(* IEC 61131-3 sources: stonehenge-public/apps/core/stonehenge-safety-plc/pous/programs, 1 file *)

(* ---- main.st ---- *)
PROGRAM main
  VAR
    SafetyGlobal : FB_GlobalSafety;
    Gun1Safety : FB_GunSafety;
    Gun2Safety : FB_GunSafety;
    Gun3Safety : FB_GunSafety;
    Gun4Safety : FB_GunSafety;
    Gun5Safety : FB_GunSafety;
    Gun6Safety : FB_GunSafety;
    Gun7Safety : FB_GunSafety;
    Gun8Safety : FB_GunSafety;
    CONTROL_VERSION_REQUEST : INT AT %MW0 := 0;
    GLOBAL_ENABLE : INT AT %MW1 := 0;
    EMERGENCY_STOP : INT AT %MW2 := 0;
    GLOBAL_MAINTENANCE_MODE : INT AT %MW3 := 0;
    SAFETY_RESET_REQUEST : INT AT %MW4 := 0;
    TEST_FAULT_REQUEST : INT AT %MW5 := 0;
    INPUT_RESERVED_6 : INT AT %MW6 := 0;
    INPUT_RESERVED_7 : INT AT %MW7 := 0;
    GUN1_ENABLED : INT AT %MW16 := 0;
    GUN1_MAINTENANCE_INHIBIT : INT AT %MW17 := 0;
    GUN1_EXTERNAL_INHIBIT : INT AT %MW18 := 0;
    GUN1_INPUT_RESERVED : INT AT %MW19 := 0;
    GUN2_ENABLED : INT AT %MW20 := 0;
    GUN2_MAINTENANCE_INHIBIT : INT AT %MW21 := 0;
    GUN2_EXTERNAL_INHIBIT : INT AT %MW22 := 0;
    GUN2_INPUT_RESERVED : INT AT %MW23 := 0;
    GUN3_ENABLED : INT AT %MW24 := 0;
    GUN3_MAINTENANCE_INHIBIT : INT AT %MW25 := 0;
    GUN3_EXTERNAL_INHIBIT : INT AT %MW26 := 0;
    GUN3_INPUT_RESERVED : INT AT %MW27 := 0;
    GUN4_ENABLED : INT AT %MW28 := 0;
    GUN4_MAINTENANCE_INHIBIT : INT AT %MW29 := 0;
    GUN4_EXTERNAL_INHIBIT : INT AT %MW30 := 0;
    GUN4_INPUT_RESERVED : INT AT %MW31 := 0;
    GUN5_ENABLED : INT AT %MW32 := 0;
    GUN5_MAINTENANCE_INHIBIT : INT AT %MW33 := 0;
    GUN5_EXTERNAL_INHIBIT : INT AT %MW34 := 0;
    GUN5_INPUT_RESERVED : INT AT %MW35 := 0;
    GUN6_ENABLED : INT AT %MW36 := 0;
    GUN6_MAINTENANCE_INHIBIT : INT AT %MW37 := 0;
    GUN6_EXTERNAL_INHIBIT : INT AT %MW38 := 0;
    GUN6_INPUT_RESERVED : INT AT %MW39 := 0;
    GUN7_ENABLED : INT AT %MW40 := 0;
    GUN7_MAINTENANCE_INHIBIT : INT AT %MW41 := 0;
    GUN7_EXTERNAL_INHIBIT : INT AT %MW42 := 0;
    GUN7_INPUT_RESERVED : INT AT %MW43 := 0;
    GUN8_ENABLED : INT AT %MW44 := 0;
    GUN8_MAINTENANCE_INHIBIT : INT AT %MW45 := 0;
    GUN8_EXTERNAL_INHIBIT : INT AT %MW46 := 0;
    GUN8_INPUT_RESERVED : INT AT %MW47 := 0;
    SAFETY_SCHEMA_VERSION : INT AT %QW0 := 0;
    SAFETY_HEARTBEAT_COUNTER : INT AT %QW1 := 0;
    SAFETY_STATE : INT AT %QW2 := 0;
    SAFETY_READY : INT AT %QW3 := 0;
    GLOBAL_FIRE_PERMISSIVE : INT AT %QW4 := 0;
    GLOBAL_INHIBIT_ACTIVE : INT AT %QW5 := 0;
    GLOBAL_INHIBIT_REASON : INT AT %QW6 := 0;
    SAFETY_FAULT_ACTIVE : INT AT %QW7 := 0;
    SAFETY_FAULT_CODE : INT AT %QW8 := 0;
    RESET_REQUIRED : INT AT %QW9 := 0;
    EMERGENCY_STOP_ACTIVE : INT AT %QW10 := 0;
    MAINTENANCE_MODE_ACTIVE : INT AT %QW11 := 0;
    STATUS_RESERVED_12 : INT AT %QW12 := 0;
    STATUS_RESERVED_13 : INT AT %QW13 := 0;
    STATUS_RESERVED_14 : INT AT %QW14 := 0;
    STATUS_RESERVED_15 : INT AT %QW15 := 0;
    GUN1_FIRE_PERMISSIVE : INT AT %QW16 := 0;
    GUN1_INHIBIT_ACTIVE : INT AT %QW17 := 0;
    GUN1_INHIBIT_REASON : INT AT %QW18 := 0;
    GUN1_ENABLED_STATUS : INT AT %QW19 := 0;
    GUN1_MAINTENANCE_INHIBIT_STATUS : INT AT %QW20 := 0;
    GUN1_EXTERNAL_INHIBIT_STATUS : INT AT %QW21 := 0;
    GUN1_STATUS_RESERVED_A : INT AT %QW22 := 0;
    GUN1_STATUS_RESERVED_B : INT AT %QW23 := 0;
    GUN2_FIRE_PERMISSIVE : INT AT %QW24 := 0;
    GUN2_INHIBIT_ACTIVE : INT AT %QW25 := 0;
    GUN2_INHIBIT_REASON : INT AT %QW26 := 0;
    GUN2_ENABLED_STATUS : INT AT %QW27 := 0;
    GUN2_MAINTENANCE_INHIBIT_STATUS : INT AT %QW28 := 0;
    GUN2_EXTERNAL_INHIBIT_STATUS : INT AT %QW29 := 0;
    GUN2_STATUS_RESERVED_A : INT AT %QW30 := 0;
    GUN2_STATUS_RESERVED_B : INT AT %QW31 := 0;
    GUN3_FIRE_PERMISSIVE : INT AT %QW32 := 0;
    GUN3_INHIBIT_ACTIVE : INT AT %QW33 := 0;
    GUN3_INHIBIT_REASON : INT AT %QW34 := 0;
    GUN3_ENABLED_STATUS : INT AT %QW35 := 0;
    GUN3_MAINTENANCE_INHIBIT_STATUS : INT AT %QW36 := 0;
    GUN3_EXTERNAL_INHIBIT_STATUS : INT AT %QW37 := 0;
    GUN3_STATUS_RESERVED_A : INT AT %QW38 := 0;
    GUN3_STATUS_RESERVED_B : INT AT %QW39 := 0;
    GUN4_FIRE_PERMISSIVE : INT AT %QW40 := 0;
    GUN4_INHIBIT_ACTIVE : INT AT %QW41 := 0;
    GUN4_INHIBIT_REASON : INT AT %QW42 := 0;
    GUN4_ENABLED_STATUS : INT AT %QW43 := 0;
    GUN4_MAINTENANCE_INHIBIT_STATUS : INT AT %QW44 := 0;
    GUN4_EXTERNAL_INHIBIT_STATUS : INT AT %QW45 := 0;
    GUN4_STATUS_RESERVED_A : INT AT %QW46 := 0;
    GUN4_STATUS_RESERVED_B : INT AT %QW47 := 0;
    GUN5_FIRE_PERMISSIVE : INT AT %QW48 := 0;
    GUN5_INHIBIT_ACTIVE : INT AT %QW49 := 0;
    GUN5_INHIBIT_REASON : INT AT %QW50 := 0;
    GUN5_ENABLED_STATUS : INT AT %QW51 := 0;
    GUN5_MAINTENANCE_INHIBIT_STATUS : INT AT %QW52 := 0;
    GUN5_EXTERNAL_INHIBIT_STATUS : INT AT %QW53 := 0;
    GUN5_STATUS_RESERVED_A : INT AT %QW54 := 0;
    GUN5_STATUS_RESERVED_B : INT AT %QW55 := 0;
    GUN6_FIRE_PERMISSIVE : INT AT %QW56 := 0;
    GUN6_INHIBIT_ACTIVE : INT AT %QW57 := 0;
    GUN6_INHIBIT_REASON : INT AT %QW58 := 0;
    GUN6_ENABLED_STATUS : INT AT %QW59 := 0;
    GUN6_MAINTENANCE_INHIBIT_STATUS : INT AT %QW60 := 0;
    GUN6_EXTERNAL_INHIBIT_STATUS : INT AT %QW61 := 0;
    GUN6_STATUS_RESERVED_A : INT AT %QW62 := 0;
    GUN6_STATUS_RESERVED_B : INT AT %QW63 := 0;
    GUN7_FIRE_PERMISSIVE : INT AT %QW64 := 0;
    GUN7_INHIBIT_ACTIVE : INT AT %QW65 := 0;
    GUN7_INHIBIT_REASON : INT AT %QW66 := 0;
    GUN7_ENABLED_STATUS : INT AT %QW67 := 0;
    GUN7_MAINTENANCE_INHIBIT_STATUS : INT AT %QW68 := 0;
    GUN7_EXTERNAL_INHIBIT_STATUS : INT AT %QW69 := 0;
    GUN7_STATUS_RESERVED_A : INT AT %QW70 := 0;
    GUN7_STATUS_RESERVED_B : INT AT %QW71 := 0;
    GUN8_FIRE_PERMISSIVE : INT AT %QW72 := 0;
    GUN8_INHIBIT_ACTIVE : INT AT %QW73 := 0;
    GUN8_INHIBIT_REASON : INT AT %QW74 := 0;
    GUN8_ENABLED_STATUS : INT AT %QW75 := 0;
    GUN8_MAINTENANCE_INHIBIT_STATUS : INT AT %QW76 := 0;
    GUN8_EXTERNAL_INHIBIT_STATUS : INT AT %QW77 := 0;
    GUN8_STATUS_RESERVED_A : INT AT %QW78 := 0;
    GUN8_STATUS_RESERVED_B : INT AT %QW79 := 0;
  END_VAR

SafetyGlobal(
    global_enable := GLOBAL_ENABLE <> 0,
    emergency_stop := EMERGENCY_STOP <> 0,
    global_maintenance_mode := GLOBAL_MAINTENANCE_MODE <> 0,
    safety_reset_request := SAFETY_RESET_REQUEST <> 0,
    test_fault_request := TEST_FAULT_REQUEST <> 0
);

Gun1Safety(global_fire_permissive := SafetyGlobal.global_fire_permissive, global_fault_active := SafetyGlobal.safety_fault_active, reset_required := SafetyGlobal.reset_required, gun_enabled := GUN1_ENABLED <> 0, gun_maintenance_inhibit := GUN1_MAINTENANCE_INHIBIT <> 0, gun_external_inhibit := GUN1_EXTERNAL_INHIBIT <> 0);
Gun2Safety(global_fire_permissive := SafetyGlobal.global_fire_permissive, global_fault_active := SafetyGlobal.safety_fault_active, reset_required := SafetyGlobal.reset_required, gun_enabled := GUN2_ENABLED <> 0, gun_maintenance_inhibit := GUN2_MAINTENANCE_INHIBIT <> 0, gun_external_inhibit := GUN2_EXTERNAL_INHIBIT <> 0);
Gun3Safety(global_fire_permissive := SafetyGlobal.global_fire_permissive, global_fault_active := SafetyGlobal.safety_fault_active, reset_required := SafetyGlobal.reset_required, gun_enabled := GUN3_ENABLED <> 0, gun_maintenance_inhibit := GUN3_MAINTENANCE_INHIBIT <> 0, gun_external_inhibit := GUN3_EXTERNAL_INHIBIT <> 0);
Gun4Safety(global_fire_permissive := SafetyGlobal.global_fire_permissive, global_fault_active := SafetyGlobal.safety_fault_active, reset_required := SafetyGlobal.reset_required, gun_enabled := GUN4_ENABLED <> 0, gun_maintenance_inhibit := GUN4_MAINTENANCE_INHIBIT <> 0, gun_external_inhibit := GUN4_EXTERNAL_INHIBIT <> 0);
Gun5Safety(global_fire_permissive := SafetyGlobal.global_fire_permissive, global_fault_active := SafetyGlobal.safety_fault_active, reset_required := SafetyGlobal.reset_required, gun_enabled := GUN5_ENABLED <> 0, gun_maintenance_inhibit := GUN5_MAINTENANCE_INHIBIT <> 0, gun_external_inhibit := GUN5_EXTERNAL_INHIBIT <> 0);
Gun6Safety(global_fire_permissive := SafetyGlobal.global_fire_permissive, global_fault_active := SafetyGlobal.safety_fault_active, reset_required := SafetyGlobal.reset_required, gun_enabled := GUN6_ENABLED <> 0, gun_maintenance_inhibit := GUN6_MAINTENANCE_INHIBIT <> 0, gun_external_inhibit := GUN6_EXTERNAL_INHIBIT <> 0);
Gun7Safety(global_fire_permissive := SafetyGlobal.global_fire_permissive, global_fault_active := SafetyGlobal.safety_fault_active, reset_required := SafetyGlobal.reset_required, gun_enabled := GUN7_ENABLED <> 0, gun_maintenance_inhibit := GUN7_MAINTENANCE_INHIBIT <> 0, gun_external_inhibit := GUN7_EXTERNAL_INHIBIT <> 0);
Gun8Safety(global_fire_permissive := SafetyGlobal.global_fire_permissive, global_fault_active := SafetyGlobal.safety_fault_active, reset_required := SafetyGlobal.reset_required, gun_enabled := GUN8_ENABLED <> 0, gun_maintenance_inhibit := GUN8_MAINTENANCE_INHIBIT <> 0, gun_external_inhibit := GUN8_EXTERNAL_INHIBIT <> 0);

SAFETY_SCHEMA_VERSION := SafetyGlobal.schema_version;
SAFETY_HEARTBEAT_COUNTER := SafetyGlobal.heartbeat_counter;
SAFETY_STATE := SafetyGlobal.safety_state;
IF SafetyGlobal.safety_ready THEN SAFETY_READY := 1; ELSE SAFETY_READY := 0; END_IF;
IF SafetyGlobal.global_fire_permissive THEN GLOBAL_FIRE_PERMISSIVE := 1; ELSE GLOBAL_FIRE_PERMISSIVE := 0; END_IF;
IF SafetyGlobal.global_inhibit_active THEN GLOBAL_INHIBIT_ACTIVE := 1; ELSE GLOBAL_INHIBIT_ACTIVE := 0; END_IF;
GLOBAL_INHIBIT_REASON := SafetyGlobal.global_inhibit_reason;
IF SafetyGlobal.safety_fault_active THEN SAFETY_FAULT_ACTIVE := 1; ELSE SAFETY_FAULT_ACTIVE := 0; END_IF;
SAFETY_FAULT_CODE := SafetyGlobal.safety_fault_code;
IF SafetyGlobal.reset_required THEN RESET_REQUIRED := 1; ELSE RESET_REQUIRED := 0; END_IF;
IF SafetyGlobal.emergency_stop_active THEN EMERGENCY_STOP_ACTIVE := 1; ELSE EMERGENCY_STOP_ACTIVE := 0; END_IF;
IF SafetyGlobal.maintenance_mode_active THEN MAINTENANCE_MODE_ACTIVE := 1; ELSE MAINTENANCE_MODE_ACTIVE := 0; END_IF;
STATUS_RESERVED_12 := 0;
STATUS_RESERVED_13 := 0;
STATUS_RESERVED_14 := 0;
STATUS_RESERVED_15 := 0;

IF Gun1Safety.fire_permissive THEN GUN1_FIRE_PERMISSIVE := 1; ELSE GUN1_FIRE_PERMISSIVE := 0; END_IF;
IF Gun1Safety.inhibit_active THEN GUN1_INHIBIT_ACTIVE := 1; ELSE GUN1_INHIBIT_ACTIVE := 0; END_IF;
GUN1_INHIBIT_REASON := Gun1Safety.inhibit_reason;
IF GUN1_ENABLED <> 0 THEN GUN1_ENABLED_STATUS := 1; ELSE GUN1_ENABLED_STATUS := 0; END_IF;
IF GUN1_MAINTENANCE_INHIBIT <> 0 THEN GUN1_MAINTENANCE_INHIBIT_STATUS := 1; ELSE GUN1_MAINTENANCE_INHIBIT_STATUS := 0; END_IF;
IF GUN1_EXTERNAL_INHIBIT <> 0 THEN GUN1_EXTERNAL_INHIBIT_STATUS := 1; ELSE GUN1_EXTERNAL_INHIBIT_STATUS := 0; END_IF;
GUN1_STATUS_RESERVED_A := 0;
GUN1_STATUS_RESERVED_B := 0;

IF Gun2Safety.fire_permissive THEN GUN2_FIRE_PERMISSIVE := 1; ELSE GUN2_FIRE_PERMISSIVE := 0; END_IF;
IF Gun2Safety.inhibit_active THEN GUN2_INHIBIT_ACTIVE := 1; ELSE GUN2_INHIBIT_ACTIVE := 0; END_IF;
GUN2_INHIBIT_REASON := Gun2Safety.inhibit_reason;
IF GUN2_ENABLED <> 0 THEN GUN2_ENABLED_STATUS := 1; ELSE GUN2_ENABLED_STATUS := 0; END_IF;
IF GUN2_MAINTENANCE_INHIBIT <> 0 THEN GUN2_MAINTENANCE_INHIBIT_STATUS := 1; ELSE GUN2_MAINTENANCE_INHIBIT_STATUS := 0; END_IF;
IF GUN2_EXTERNAL_INHIBIT <> 0 THEN GUN2_EXTERNAL_INHIBIT_STATUS := 1; ELSE GUN2_EXTERNAL_INHIBIT_STATUS := 0; END_IF;
GUN2_STATUS_RESERVED_A := 0;
GUN2_STATUS_RESERVED_B := 0;

IF Gun3Safety.fire_permissive THEN GUN3_FIRE_PERMISSIVE := 1; ELSE GUN3_FIRE_PERMISSIVE := 0; END_IF;
IF Gun3Safety.inhibit_active THEN GUN3_INHIBIT_ACTIVE := 1; ELSE GUN3_INHIBIT_ACTIVE := 0; END_IF;
GUN3_INHIBIT_REASON := Gun3Safety.inhibit_reason;
IF GUN3_ENABLED <> 0 THEN GUN3_ENABLED_STATUS := 1; ELSE GUN3_ENABLED_STATUS := 0; END_IF;
IF GUN3_MAINTENANCE_INHIBIT <> 0 THEN GUN3_MAINTENANCE_INHIBIT_STATUS := 1; ELSE GUN3_MAINTENANCE_INHIBIT_STATUS := 0; END_IF;
IF GUN3_EXTERNAL_INHIBIT <> 0 THEN GUN3_EXTERNAL_INHIBIT_STATUS := 1; ELSE GUN3_EXTERNAL_INHIBIT_STATUS := 0; END_IF;
GUN3_STATUS_RESERVED_A := 0;
GUN3_STATUS_RESERVED_B := 0;

IF Gun4Safety.fire_permissive THEN GUN4_FIRE_PERMISSIVE := 1; ELSE GUN4_FIRE_PERMISSIVE := 0; END_IF;
IF Gun4Safety.inhibit_active THEN GUN4_INHIBIT_ACTIVE := 1; ELSE GUN4_INHIBIT_ACTIVE := 0; END_IF;
GUN4_INHIBIT_REASON := Gun4Safety.inhibit_reason;
IF GUN4_ENABLED <> 0 THEN GUN4_ENABLED_STATUS := 1; ELSE GUN4_ENABLED_STATUS := 0; END_IF;
IF GUN4_MAINTENANCE_INHIBIT <> 0 THEN GUN4_MAINTENANCE_INHIBIT_STATUS := 1; ELSE GUN4_MAINTENANCE_INHIBIT_STATUS := 0; END_IF;
IF GUN4_EXTERNAL_INHIBIT <> 0 THEN GUN4_EXTERNAL_INHIBIT_STATUS := 1; ELSE GUN4_EXTERNAL_INHIBIT_STATUS := 0; END_IF;
GUN4_STATUS_RESERVED_A := 0;
GUN4_STATUS_RESERVED_B := 0;

IF Gun5Safety.fire_permissive THEN GUN5_FIRE_PERMISSIVE := 1; ELSE GUN5_FIRE_PERMISSIVE := 0; END_IF;
IF Gun5Safety.inhibit_active THEN GUN5_INHIBIT_ACTIVE := 1; ELSE GUN5_INHIBIT_ACTIVE := 0; END_IF;
GUN5_INHIBIT_REASON := Gun5Safety.inhibit_reason;
IF GUN5_ENABLED <> 0 THEN GUN5_ENABLED_STATUS := 1; ELSE GUN5_ENABLED_STATUS := 0; END_IF;
IF GUN5_MAINTENANCE_INHIBIT <> 0 THEN GUN5_MAINTENANCE_INHIBIT_STATUS := 1; ELSE GUN5_MAINTENANCE_INHIBIT_STATUS := 0; END_IF;
IF GUN5_EXTERNAL_INHIBIT <> 0 THEN GUN5_EXTERNAL_INHIBIT_STATUS := 1; ELSE GUN5_EXTERNAL_INHIBIT_STATUS := 0; END_IF;
GUN5_STATUS_RESERVED_A := 0;
GUN5_STATUS_RESERVED_B := 0;

IF Gun6Safety.fire_permissive THEN GUN6_FIRE_PERMISSIVE := 1; ELSE GUN6_FIRE_PERMISSIVE := 0; END_IF;
IF Gun6Safety.inhibit_active THEN GUN6_INHIBIT_ACTIVE := 1; ELSE GUN6_INHIBIT_ACTIVE := 0; END_IF;
GUN6_INHIBIT_REASON := Gun6Safety.inhibit_reason;
IF GUN6_ENABLED <> 0 THEN GUN6_ENABLED_STATUS := 1; ELSE GUN6_ENABLED_STATUS := 0; END_IF;
IF GUN6_MAINTENANCE_INHIBIT <> 0 THEN GUN6_MAINTENANCE_INHIBIT_STATUS := 1; ELSE GUN6_MAINTENANCE_INHIBIT_STATUS := 0; END_IF;
IF GUN6_EXTERNAL_INHIBIT <> 0 THEN GUN6_EXTERNAL_INHIBIT_STATUS := 1; ELSE GUN6_EXTERNAL_INHIBIT_STATUS := 0; END_IF;
GUN6_STATUS_RESERVED_A := 0;
GUN6_STATUS_RESERVED_B := 0;

IF Gun7Safety.fire_permissive THEN GUN7_FIRE_PERMISSIVE := 1; ELSE GUN7_FIRE_PERMISSIVE := 0; END_IF;
IF Gun7Safety.inhibit_active THEN GUN7_INHIBIT_ACTIVE := 1; ELSE GUN7_INHIBIT_ACTIVE := 0; END_IF;
GUN7_INHIBIT_REASON := Gun7Safety.inhibit_reason;
IF GUN7_ENABLED <> 0 THEN GUN7_ENABLED_STATUS := 1; ELSE GUN7_ENABLED_STATUS := 0; END_IF;
IF GUN7_MAINTENANCE_INHIBIT <> 0 THEN GUN7_MAINTENANCE_INHIBIT_STATUS := 1; ELSE GUN7_MAINTENANCE_INHIBIT_STATUS := 0; END_IF;
IF GUN7_EXTERNAL_INHIBIT <> 0 THEN GUN7_EXTERNAL_INHIBIT_STATUS := 1; ELSE GUN7_EXTERNAL_INHIBIT_STATUS := 0; END_IF;
GUN7_STATUS_RESERVED_A := 0;
GUN7_STATUS_RESERVED_B := 0;

IF Gun8Safety.fire_permissive THEN GUN8_FIRE_PERMISSIVE := 1; ELSE GUN8_FIRE_PERMISSIVE := 0; END_IF;
IF Gun8Safety.inhibit_active THEN GUN8_INHIBIT_ACTIVE := 1; ELSE GUN8_INHIBIT_ACTIVE := 0; END_IF;
GUN8_INHIBIT_REASON := Gun8Safety.inhibit_reason;
IF GUN8_ENABLED <> 0 THEN GUN8_ENABLED_STATUS := 1; ELSE GUN8_ENABLED_STATUS := 0; END_IF;
IF GUN8_MAINTENANCE_INHIBIT <> 0 THEN GUN8_MAINTENANCE_INHIBIT_STATUS := 1; ELSE GUN8_MAINTENANCE_INHIBIT_STATUS := 0; END_IF;
IF GUN8_EXTERNAL_INHIBIT <> 0 THEN GUN8_EXTERNAL_INHIBIT_STATUS := 1; ELSE GUN8_EXTERNAL_INHIBIT_STATUS := 0; END_IF;
GUN8_STATUS_RESERVED_A := 0;
GUN8_STATUS_RESERVED_B := 0;

END_PROGRAM
